Fanuc KAREL source: kt00724.KL

-- PROVISIONAL review KL for V1013-1; original PC SHA256 f602626a528b3946fc52f0cd543168ed1a17379510c151adf95b909ea8b89e79
-- Incomplete behavior may be omitted. Consult companion uncertainty JSON. Do not deploy.
PROGRAM KT00724
%NOLOCKGROUP
VAR
  OUT : BOOLEAN
-- UNRESOLVED_DECL P1 type=000199
-- UNRESOLVED_DECL P2 type=000199
BEGIN
  -- UNRESOLVED_PC offsets 5-20; opcodes 22,63,23
  -- UNRESOLVED_PC offsets 25-29; opcodes 7F
END KT00724
